(*
SPDX-FileCopyrightText: © 2026 Oleksandr Tiutyk <trofimich@gmail.com>
SPDX-License-Identifier: MIT
License: https://opensource.org/license/mit
*)

(*!
<summary>Test workflow instance containing named variables for the comprehensive workflow scenario test.</summary>
*)

{attribute 'no_explicit_call' := 'do not call this function block directly'}
{attribute 'enable_dynamic_creation'}
FUNCTION_BLOCK ComprehensiveTestWorkflow EXTENDS TOF_Workflow.Workflow
VAR_INPUT
	SensorFeedPart : BOOL;
	SensorVacuumOk : BOOL;
	SensorInspectionOk : BOOL;
	BatchTarget : INT;
	ProducedCount : INT;
	RejectCount : INT;
	ErrorHandled : BOOL;
END_VAR
VAR_STAT
	//! <summary>Concrete test workflow name available during inherited initialization.</summary>
	_TestWorkflowClassName : STRING := __POUNAME();
END_VAR

METHOD PROTECTED InitializeVariables
BindPlcVariable(name := 'BatchTarget', plcVariable := BatchTarget);
BindPlcVariable(name := 'ProducedCount', plcVariable := ProducedCount);
BindPlcVariable(name := 'RejectCount', plcVariable := RejectCount);
BindPlcVariable(name := 'SensorFeedPart', plcVariable := SensorFeedPart);
BindPlcVariable(name := 'SensorVacuumOk', plcVariable := SensorVacuumOk);
BindPlcVariable(name := 'SensorInspectionOk', plcVariable := SensorInspectionOk);
BindPlcVariable(name := 'ErrorHandled', plcVariable := ErrorHandled);
END_METHOD

{attribute 'monitoring' := 'call'}
PROPERTY NamespaceName : REFERENCE TO STRING
GET
NamespaceName REF= CurrentNamespace.Name;
END_GET
END_PROPERTY

METHOD PROTECTED OnRootActivityRequestReset
VAR_OUTPUT
	abortRequest : BOOL;
END_VAR
ProducedCount := 0;
RejectCount := 0;
ErrorHandled := FALSE;
END_METHOD

{attribute 'monitoring' := 'call'}
PROPERTY SelfSize : ULINT
GET
SelfSize := XSIZEOF(THIS^);
END_GET
END_PROPERTY

(*!
<summary>Returns the concrete test workflow name from initialized static storage.</summary>
*)
{attribute 'monitoring' := 'call'}
PROPERTY ClassName : REFERENCE TO STRING
GET
ClassName REF= _TestWorkflowClassName;
END_GET
END_PROPERTY

END_FUNCTION_BLOCK

(* stored: Version 1.1.0.1, ProductVersion 3.1.4026.21
   POU ComprehensiveTestWorkflow: Id {f68cdb29-f402-4a3c-a63d-1d66373aec54}, SpecialFunc None
   Folder Overriden members: Id {e4c1214b-c5de-4258-be55-74a6472c32e0}
   Method InitializeVariables: Id {ca266811-7478-4488-af0f-64a400c7b49b}
   Property NamespaceName: Id {0883b169-afc6-4537-86f5-2fd46e0faffe}
   Get Get: Id {142455da-6cd3-477b-ac63-8ab44d5d32bc}
   Method OnRootActivityRequestReset: Id {40bfb420-e972-4486-a912-6873773be130}
   Property SelfSize: Id {0a9b2890-9932-44fe-a7d7-72edc5b13608}
   Get Get: Id {a533cfa1-ac99-4f9f-a92d-a5810418a3c1}
   Property ClassName: Id {84492f4a-0290-4c01-9eb5-0e24af66383a}
   Get Get: Id {85400a5e-c5c7-4c22-a6f8-489fa5b4b293} *)
